FUNCTION_BLOCK EV_LinearAxis (* Names the equipment's two channels, and unpacks its state channel into named values (its inputs and who holds it) for a skill. Technical: Names LinearAxis's channels; typed view of its state channel (inputs and holder) *)
  (* Standard: 61499-2 *)
  (* Version 0.1, 2026-09-28, Project contributors, AAU Smart Production Lab *)
  PACKAGE capping;
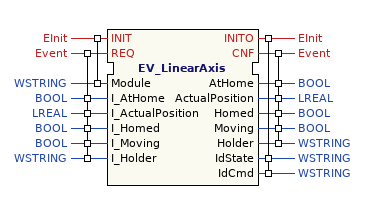
  EVENT_INPUT
    INIT : EInit WITH Module; (* Name the equipment's channels *)
    REQ WITH I_AtHome, I_ActualPosition, I_Homed, I_Moving, I_Holder; (* The equipment's state arrived *)
  END_EVENT
  EVENT_OUTPUT
    INITO : EInit WITH IdState, IdCmd; (* IdState and IdCmd are set *)
    CNF WITH AtHome, ActualPosition, Homed, Moving, Holder; (* The values below are updated *)
  END_EVENT
  VAR_INPUT
    Module : WSTRING; (* The module's name; its local channels are named after it (loc[<Module>/...]) *)
    I_AtHome : BOOL; (* AtHome as read or received *)
    I_ActualPosition : LREAL; (* ActualPosition as read or received *)
    I_Homed : BOOL; (* Homed as read or received *)
    I_Moving : BOOL; (* Moving as read or received *)
    I_Holder : WSTRING; (* Holder as read or received *)
  END_VAR
  VAR_OUTPUT
    AtHome : BOOL; (* LinearAxis: AtHome, an input *)
    ActualPosition : LREAL; (* LinearAxis: ActualPosition (mm), worked out by the equipment *)
    Homed : BOOL; (* LinearAxis: Homed, worked out by the equipment *)
    Moving : BOOL; (* LinearAxis: Moving, worked out by the equipment *)
    Holder : WSTRING; (* Who holds the equipment (empty: free) *)
    IdState : WSTRING; (* Local channel of the equipment's state *)
    IdCmd : WSTRING; (* Local channel of the equipment's commands *)
  END_VAR
  EC_STATES
    INIT : INIT -> INITO;
    REQ : REQ -> CNF;
  END_STATES
  ALGORITHM INIT IN ST:
IdState := CONCAT(CONCAT("loc[", Module), "/LinearAxis/state]");
IdCmd := CONCAT(CONCAT("loc[", Module), "/LinearAxis/cmd]");
  END_ALGORITHM
  ALGORITHM REQ IN ST:
AtHome := I_AtHome;
ActualPosition := I_ActualPosition;
Homed := I_Homed;
Moving := I_Moving;
Holder := I_Holder;
  END_ALGORITHM
END_FUNCTION_BLOCK
